FUNCTION_BLOCK FB_Maschine IMPLEMENTS I_Maschine
VAR
	_zustand : E_Zustand := E_Zustand.Aus;
	_notaus : BOOL := FALSE;
END_VAR

METHOD Start
IF NOT _notaus THEN
	_zustand := E_Zustand.Bereit;
END_IF
END_METHOD

METHOD Stop
_zustand := E_Zustand.Aus;
END_METHOD

METHOD NotausAusloesen
_notaus := TRUE;
_zustand := E_Zustand.Notaus;
END_METHOD

METHOD NotausZuruecksetzen
_notaus := FALSE;
_zustand := E_Zustand.Bereit;
END_METHOD

PROPERTY Zustand : E_Zustand
END_PROPERTY

END_FUNCTION_BLOCK

(* stored: Version 1.1.0.1, ProductVersion 3.1.4024.32
   POU FB_Maschine: Id {F7C8490A-1B2C-4738-594A-C5D6E7F8091A}, SpecialFunc None
   Method Start: Id {5D904F61-7283-4E9F-A01B-2C3D4E5F6071}
   Method Stop: Id {6EA15072-8394-4FA0-B12C-3D4E5F607182}
   Method NotausAusloesen: Id {7FB26183-94A5-40B1-C23D-4E5F60718293}
   Method NotausZuruecksetzen: Id {80C37294-A5B6-41C2-D34E-5F60718293A4}
   Property Zustand: Id {91D483A5-B6C7-42D3-E45F-60718293A4B5} *)
